DATA_BLOCK "FRK_EventDeliveryView"
{ S7_Optimized_Access := 'TRUE' }
VERSION : 0.1
NON_RETAIN
VAR
    Count {ExternalWritable := 'False'} : Int := 1;
    Rows {ExternalWritable := 'False'} : Array[1..1] of "FRK_DeliveryView";
END_VAR
BEGIN
END_DATA_BLOCK
